Universal Robots PolyScope program: Put_into_box_E-series_UR10.urp

Program  (createdIn=3.0.0.0 lastSavedIn=5.0.3.30563)
Robot Program (runOnlyOnce=true speed=0 acceleration=0 useActiveTCP=false positionType=CartesianPose) feature=Base
  Set NoAction (payload=0 tcpAsCog=true)
  MoveJ speed 50 deg/s, acceleration 100 deg/s^2 (useActiveTCP=false positionType=JointAngles)
    Waypoint Home: TCP in base x=-0.004 y=-290.7 z=1484.8 mm, rx=0 ry=2.2214 rz=-2.2214 rad; joints [0.001, -90, 0, -90, -0.001, 0.001] deg
    Waypoint End: TCP in base x=-147.934 y=57.6 z=121.475 mm, rx=0.0001 ry=-2.2214 rz=2.2214 rad; joints [180, -90, -165, -105, 180.001, 179.997] deg
